TYPE "FRK_Document_D019"
VERSION : 0.1
   STRUCT
      "SchemaVersion" {ExternalAccessible := 'False'; ExternalVisible := 'False'; ExternalWritable := 'False'} : UInt;
      "Scope" {ExternalAccessible := 'False'; ExternalVisible := 'False'; ExternalWritable := 'False'} : String[80];
      "Image" {ExternalAccessible := 'False'; ExternalVisible := 'False'; ExternalWritable := 'False'} : "FRK_ClassPolicyImage";
   END_STRUCT;
END_TYPE
